Fanuc KAREL source: KD00051.KL

PROGRAM KD00051
%NOLOCKGROUP
%DEFGROUP = 1
VAR
  I: INTEGER
  J: INTEGER
  B: BOOLEAN
  R: REAL
  S: STRING[80]
  P: POSITION
BEGIN
  MOVE NEAR P BY 10.0
END KD00051
